(* IEC 61131-3 sources: trust-platform/crates/trust-runtime/tests/fixtures/oscat/core/src/05_mathematics, 1 file *)

(* ---- tests.st ---- *)
TEST_PROGRAM oscat_math_helpers_behave
ASSERT_TRUE(IN := OSCAT_BASIC_Constants());
ASSERT_EQUAL(EXPECTED := DINT#3, ACTUAL := FLOOR2(X := REAL#3.14));
ASSERT_EQUAL(EXPECTED := DINT#-4, ACTUAL := FLOOR2(X := REAL#-3.14));
ASSERT_NEAR(EXPECTED := REAL#0.5, ACTUAL := MODR(IN := REAL#5.5, DIVI := REAL#2.5), DELTA := REAL#0.001);
ASSERT_NEAR(EXPECTED := REAL#180.0, ACTUAL := DEG(rad := MATH.PI), DELTA := REAL#0.01);
ASSERT_NEAR(EXPECTED := MATH.PI, ACTUAL := RAD(DEG := REAL#180.0), DELTA := REAL#0.001);
ASSERT_NEAR(EXPECTED := REAL#5.0, ACTUAL := HYPOT(X := REAL#3.0, Y := REAL#4.0), DELTA := REAL#0.001);
ASSERT_NEAR(EXPECTED := REAL#1000.0, ACTUAL := EXP10(X := REAL#3.0), DELTA := REAL#0.1);
END_TEST_PROGRAM

TEST_PROGRAM oscat_extended_math_helpers_behave
ASSERT_TRUE(IN := OSCAT_BASIC_Constants());
ASSERT_NEAR(EXPECTED := REAL#0.0, ACTUAL := AGDF(X := REAL#0.0), DELTA := REAL#0.001);
ASSERT_NEAR(EXPECTED := REAL#0.0, ACTUAL := ACOSH(X := REAL#1.0), DELTA := REAL#0.001);
ASSERT_NEAR(EXPECTED := REAL#0.549306, ACTUAL := ACOTH(X := REAL#2.0), DELTA := REAL#0.001);
ASSERT_NEAR(EXPECTED := REAL#0.0, ACTUAL := ASINH(X := REAL#0.0), DELTA := REAL#0.001);
ASSERT_NEAR(EXPECTED := MATH.PI05, ACTUAL := ATAN2(Y := REAL#1.0, X := REAL#0.0), DELTA := REAL#0.001);
ASSERT_NEAR(EXPECTED := REAL#0.549306, ACTUAL := ATANH(X := REAL#0.5), DELTA := REAL#0.001);
ASSERT_NEAR(EXPECTED := REAL#0.083333, ACTUAL := BETA(X := REAL#2.0, Y := REAL#3.0), DELTA := REAL#0.01);
ASSERT_EQUAL(EXPECTED := DINT#10, ACTUAL := BINOM(N := INT#5, K := INT#2));
ASSERT_NEAR(EXPECTED := MATH.PI_INV, ACTUAL := CAUCHY(X := REAL#0.0, T := REAL#0.0, U := REAL#1.0), DELTA := REAL#0.001);
ASSERT_NEAR(EXPECTED := REAL#0.5, ACTUAL := CAUCHYCD(X := REAL#0.0, T := REAL#0.0, U := REAL#1.0), DELTA := REAL#0.001);
ASSERT_NEAR(EXPECTED := REAL#1.0, ACTUAL := COSH(X := REAL#0.0), DELTA := REAL#0.001);
ASSERT_NEAR(EXPECTED := REAL#1.313035, ACTUAL := COTH(X := REAL#1.0), DELTA := REAL#0.001);
ASSERT_NEAR(EXPECTED := REAL#0.0, ACTUAL := SINH(X := REAL#0.0), DELTA := REAL#0.001);
ASSERT_NEAR(EXPECTED := REAL#0.761594, ACTUAL := TANH(X := REAL#1.0), DELTA := REAL#0.001);
ASSERT_TRUE(IN := CMP(X := REAL#3.141516, Y := REAL#3.141517, N := INT#6));
ASSERT_FALSE(IN := CMP(X := REAL#3.141516, Y := REAL#3.141517, N := INT#7));
ASSERT_EQUAL(EXPECTED := INT#4, ACTUAL := CEIL(X := REAL#3.14));
ASSERT_EQUAL(EXPECTED := DINT#-3, ACTUAL := CEIL2(X := REAL#-3.14));
ASSERT_EQUAL(EXPECTED := INT#3, ACTUAL := FLOOR(X := REAL#3.14));
ASSERT_EQUAL(EXPECTED := DINT#-1, ACTUAL := D_TRUNC(X := REAL#-1.5));
ASSERT_NEAR(EXPECTED := REAL#0.14, ACTUAL := FRACT(X := REAL#3.14), DELTA := REAL#0.001);
ASSERT_NEAR(EXPECTED := REAL#24.0, ACTUAL := GAMMA(X := REAL#5.0), DELTA := REAL#0.01);
ASSERT_EQUAL(EXPECTED := INT#2, ACTUAL := DEC1(X := INT#0, N := INT#3));
ASSERT_TRUE(IN := DIFFER(in1 := REAL#1.0, in2 := REAL#1.2, X := REAL#0.1));
ASSERT_FALSE(IN := DIFFER(in1 := REAL#1.0, in2 := REAL#1.05, X := REAL#0.1));
ASSERT_TRUE(IN := EVEN(IN := DINT#4));
ASSERT_FALSE(IN := EVEN(IN := DINT#5));
ASSERT_EQUAL(EXPECTED := INT#0, ACTUAL := INC(INT#2, INT#2, INT#3));
ASSERT_EQUAL(EXPECTED := INT#0, ACTUAL := INC1(X := INT#2, N := INT#3));
ASSERT_EQUAL(EXPECTED := INT#3, ACTUAL := INC2(INT#5, INT#2, INT#3, INT#6));
ASSERT_NEAR(EXPECTED := REAL#0.25, ACTUAL := INV(X := REAL#4.0), DELTA := REAL#0.001);
ASSERT_NEAR(EXPECTED := REAL#3.0, ACTUAL := MAX3(IN1 := REAL#3.0, IN2 := REAL#1.0, IN3 := REAL#2.0), DELTA := REAL#0.001);
ASSERT_NEAR(EXPECTED := REAL#2.0, ACTUAL := MID3(IN1 := REAL#3.0, IN2 := REAL#1.0, IN3 := REAL#2.0), DELTA := REAL#0.001);
ASSERT_NEAR(EXPECTED := REAL#1.0, ACTUAL := MIN3(IN1 := REAL#3.0, IN2 := REAL#1.0, IN3 := REAL#2.0), DELTA := REAL#0.001);
ASSERT_NEAR(EXPECTED := REAL#10.0, ACTUAL := MUL_ADD(X := REAL#2.0, K := REAL#3.0, O := REAL#4.0), DELTA := REAL#0.001);
ASSERT_NEAR(EXPECTED := REAL#-2.5, ACTUAL := NEGX(X := REAL#2.5), DELTA := REAL#0.001);
ASSERT_EQUAL(EXPECTED := INT#-1, ACTUAL := SGN(X := REAL#-0.5));
END_TEST_PROGRAM

TEST_PROGRAM oscat_probability_and_sequence_math_helpers_behave
ASSERT_TRUE(IN := OSCAT_BASIC_Constants());
ASSERT_NEAR(EXPECTED := REAL#0.842701, ACTUAL := ERF(X := REAL#1.0), DELTA := REAL#0.002);
ASSERT_NEAR(EXPECTED := REAL#0.157299, ACTUAL := ERFC(X := REAL#1.0), DELTA := REAL#0.002);
ASSERT_NEAR(EXPECTED := REAL#8.0, ACTUAL := EXPN(X := REAL#2.0, N := INT#3), DELTA := REAL#0.001);
ASSERT_NEAR(EXPECTED := REAL#0.125, ACTUAL := EXPN(X := REAL#2.0, N := INT#-3), DELTA := REAL#0.001);
ASSERT_EQUAL(EXPECTED := DINT#120, ACTUAL := FACT(X := INT#5));
ASSERT_EQUAL(EXPECTED := DINT#55, ACTUAL := FIB(X := INT#10));
ASSERT_NEAR(EXPECTED := REAL#0.398942, ACTUAL := GAUSS(X := REAL#0.0, U := REAL#0.0, SI := REAL#1.0), DELTA := REAL#0.002);
ASSERT_NEAR(EXPECTED := REAL#0.5, ACTUAL := GAUSSCD(X := REAL#0.0, U := REAL#0.0, SI := REAL#1.0), DELTA := REAL#0.002);
ASSERT_EQUAL(EXPECTED := INT#6, ACTUAL := GCD(A := DINT#48, B := DINT#18));
ASSERT_NEAR(EXPECTED := REAL#0.0, ACTUAL := GDF(X := REAL#0.0), DELTA := REAL#0.001);
ASSERT_NEAR(EXPECTED := REAL#1.618034, ACTUAL := GOLD(X := REAL#1.0), DELTA := REAL#0.001);
END_TEST_PROGRAM

TEST_PROGRAM oscat_advanced_math_helpers_behave
VAR
    Fraction : FRACTION;
END_VAR

ASSERT_TRUE(IN := OSCAT_BASIC_Constants());
ASSERT_NEAR(EXPECTED := REAL#0.567143, ACTUAL := LAMBERT_W(X := REAL#1.0), DELTA := REAL#0.002);
ASSERT_NEAR(EXPECTED := REAL#0.313035, ACTUAL := LANGEVIN(X := REAL#1.0), DELTA := REAL#0.002);
Fraction := REAL_TO_FRAC(X := REAL#0.75, N := INT#10);
ASSERT_EQUAL(EXPECTED := INT#3, ACTUAL := Fraction.NUMERATOR);
ASSERT_EQUAL(EXPECTED := INT#4, ACTUAL := Fraction.DENOMINATOR);
ASSERT_NEAR(EXPECTED := REAL#3.1, ACTUAL := RND(X := REAL#3.19, N := INT#2), DELTA := REAL#0.001);
ASSERT_NEAR(EXPECTED := REAL#3.15, ACTUAL := ROUND(IN := REAL#3.146, N := INT#2), DELTA := REAL#0.001);
ASSERT_NEAR(EXPECTED := REAL#0.5, ACTUAL := SIGMOID(X := REAL#0.0), DELTA := REAL#0.001);
ASSERT_TRUE(IN := SIGN_I(IN := DINT#-1));
ASSERT_TRUE(IN := SIGN_R(IN := REAL#-0.1));
ASSERT_NEAR(EXPECTED := REAL#1.0, ACTUAL := SINC(X := REAL#0.0), DELTA := REAL#0.001);
ASSERT_NEAR(EXPECTED := REAL#3.0, ACTUAL := SQRTN(X := REAL#27.0, N := INT#3), DELTA := REAL#0.002);
ASSERT_NEAR(EXPECTED := REAL#1.0, ACTUAL := TANC(X := REAL#0.0), DELTA := REAL#0.001);
ASSERT_TRUE(IN := WINDOW(LOW := REAL#0.0, IN := REAL#0.5, HIGH := REAL#1.0));
ASSERT_FALSE(IN := WINDOW(LOW := REAL#0.0, IN := REAL#1.0, HIGH := REAL#1.0));
ASSERT_TRUE(IN := WINDOW2(LOW := REAL#0.0, IN := REAL#1.0, HIGH := REAL#1.0));
END_TEST_PROGRAM

TEST_PROGRAM oscat_random_math_helpers_behave
VAR
    RandomReal : REAL;
    RandomInt : INT;
    RandomDw : DWORD;
END_VAR

ASSERT_TRUE(IN := OSCAT_BASIC_Constants());
RandomReal := RDM(LAST := REAL#0.25);
ASSERT_TRUE(IN := RandomReal >= REAL#0.0);
ASSERT_TRUE(IN := RandomReal <= REAL#1.0);
RandomInt := RDM2(LAST := INT#17, LOW := INT#3, HIGH := INT#6);
ASSERT_TRUE(IN := RandomInt >= INT#3);
ASSERT_TRUE(IN := RandomInt <= INT#6);
RandomDw := RDMDW(LAST := DWORD#12345);
ASSERT_TRUE(IN := BIT_COUNT(IN := RandomDw) >= INT#0);
END_TEST_PROGRAM
